(* IEC 61131-3 sources: kns-pump-station/targets/plc210/src/POUs/FieldBus/PRG_FieldBusOut_Plc210, 2 files *)

(* ---- PRG_FieldBusOut_Plc210.decl.st ---- *)
// Назначение: полевая шина сборки ОВЕН ПЛК210, выход (MainTask, последней — после PRG_FieldOut): слово
//             управления и задание частоты ПЧ Н1…Н3 → каналы записи Modbus RTU (FC16 4x 0…1). Встроенные
//             релейные выходы DO5…DO11 привязаны к GVL_IO в дереве устройств напрямую. Массивы привязывает
//             к каналам tools_project/codesys/plc210_io.py.
// Автор:      kr0nsch
// Версия:     0.1.0
// Документ:   docs/DESIGN.md, раздел 8.4; targets/plc210/README.md
PROGRAM PRG_FieldBusOut_Plc210
VAR
    awP101Wr : ARRAY[0..GVL_ConstPlc210.MB_VFD_WR_LAST] OF WORD;     // слейв 1: FC16 4x 0…1
    awP102Wr : ARRAY[0..GVL_ConstPlc210.MB_VFD_WR_LAST] OF WORD;     // слейв 2
    awP103Wr : ARRAY[0..GVL_ConstPlc210.MB_VFD_WR_LAST] OF WORD;     // слейв 3
END_VAR

(* ---- PRG_FieldBusOut_Plc210.impl.st ---- *)
IF GVL_Sim.xSimulation THEN
    RETURN;
END_IF

awP101Wr[GVL_ConstPlc210.MB_VFD_WR_CTW] := GVL_IO.wP101_CTW;
awP101Wr[GVL_ConstPlc210.MB_VFD_WR_FREF] := UINT_TO_WORD(GVL_IO.uiP101_FREF);
awP102Wr[GVL_ConstPlc210.MB_VFD_WR_CTW] := GVL_IO.wP102_CTW;
awP102Wr[GVL_ConstPlc210.MB_VFD_WR_FREF] := UINT_TO_WORD(GVL_IO.uiP102_FREF);
awP103Wr[GVL_ConstPlc210.MB_VFD_WR_CTW] := GVL_IO.wP103_CTW;
awP103Wr[GVL_ConstPlc210.MB_VFD_WR_FREF] := UINT_TO_WORD(GVL_IO.uiP103_FREF);
